(* Logix 5000 project; controller TFF vendor 1 type 14 code 107 rev 33.11; software revision 33.04; part 27 of 38 *)
(* tags used below, declared in another part *)
   Address : DINT;   // Temp Address
   FeedPump_PID_Settings : INT;   // Index
   Index : DINT;   // Index
   TIME : DINT[2];
   AnalogOutput : AnalogOutput[25];   // Analog Output Array
   Concentration : Concentration;
   ControlLoop_FeedPump : ALIAS FOR ControlLoop[1];
   ControlLoop_FeedPumpAlarm : ALIAS FOR AlarmDeviation[1];
   ControlLoop_TIC101 : ALIAS FOR ControlLoop[7];
   DerivedData : DerivedData;   // Derived data (user input and calculated values)
   DF3PHP003 : ALIAS FOR DigitalPoint[27];
   DF48P001 : ALIAS FOR DigitalPoint[23];
   Diafiltration : Diafiltration;
   DigitalOutput : BOOL[256];   // Digital Output Array these bits are sent to output cards.
   DigitalPoint : DigitalPoint[150];   // Digital Point Array
   DP : ALIAS FOR AnalogPoint[40];
   DPAlarm : ALIAS FOR AlarmAnalog[40];
   Drive : Drive[11];   // Drives Array
   FI003 : ALIAS FOR AnalogPoint[42];
   FI101 : ALIAS FOR AnalogPoint[19];
   FI201 : ALIAS FOR AnalogPoint[2];
   FI401 : ALIAS FOR AnalogPoint[20];
   FlowPath : FlowPath[64];   // Flow Path Array
   FQ_Conc : ALIAS FOR Totalizer[0];   // Concentration Totalizer
   FQ_Diaf : ALIAS FOR Totalizer[1];   // DiafiltrationTotalizer
   LI101 : ALIAS FOR AnalogPoint[44];
   Membrane_Data : Membrane_Data;   // Membrane Data
   NWP : ALIAS FOR AnalogPoint[45];
   Options : Options;   // Options List
   PERM : ALIAS FOR AnalogPoint[46];
   Phase0 : ALIAS FOR Phase[0];   // Phase 0
   PI001 : ALIAS FOR AnalogPoint[5];
   PI101 : ALIAS FOR AnalogPoint[6];
   PI201 : ALIAS FOR AnalogPoint[7];
   PipeAnimation : PipeAnimation;   // HMI Pipe Animation Array
   SIC001 : ALIAS FOR Drive[1];
   SIC001DF : ALIAS FOR DigitalPoint[16];
   SIC002 : ALIAS FOR Drive[2];
   SIC003DF : ALIAS FOR DigitalPoint[29];
   SysControl : SysControl;   // General system status and command
   TCU101_AO : ALIAS FOR AnalogOutput[6];
   TI101 : ALIAS FOR AnalogPoint[13];
   TI201 : ALIAS FOR AnalogPoint[22];
   TIC101Control : TCUControl;
   TMP : ALIAS FOR AnalogPoint[41];
   TMPAlarm : ALIAS FOR AlarmAnalog[41];
   XV701 : ALIAS FOR Valve[17];
   XV702 : ALIAS FOR Valve[18];
(* Process, continued *)

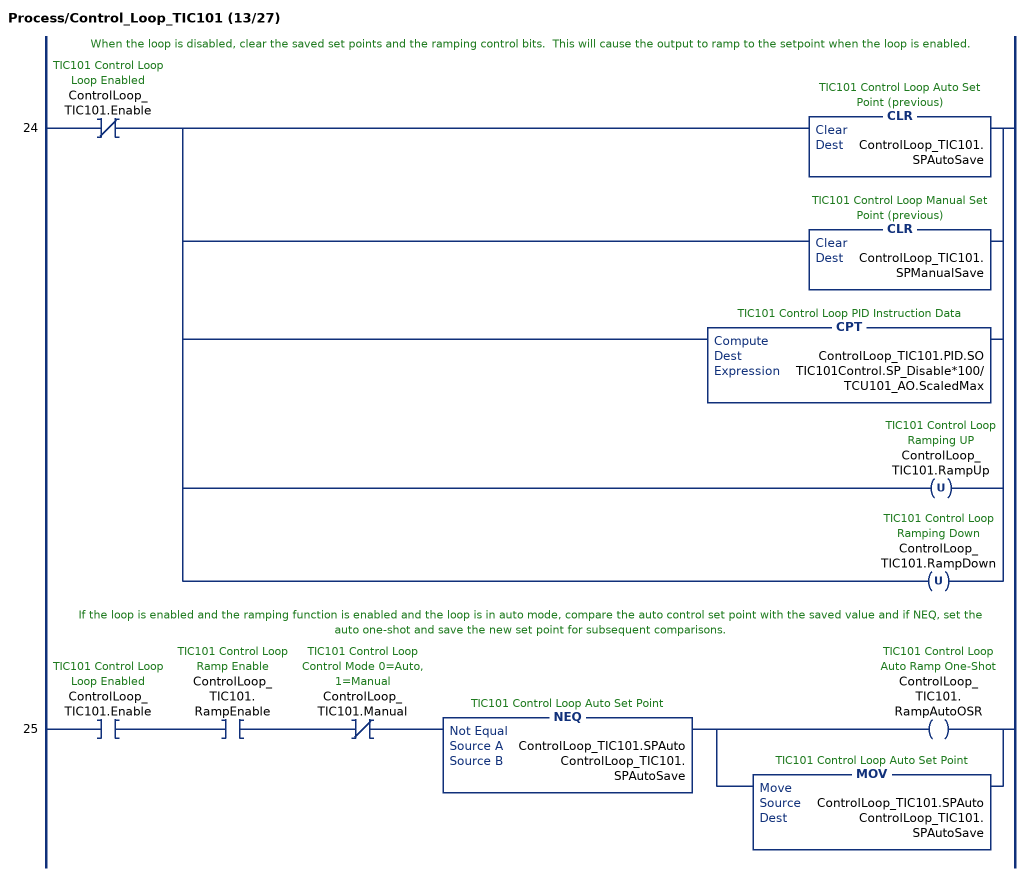
   [picture p263: Process/Control_Loop_TIC101 rungs 24-25]
   // When the loop is disabled, clear the saved set points and the ramping control bits.  This will cause the output to ramp to the setpoint when the loop is enabled.
   24: XIO(ControlLoop_TIC101.Enable)[CLR(ControlLoop_TIC101.SPAutoSave) ,CLR(ControlLoop_TIC101.SPManualSave) ,CPT(ControlLoop_TIC101.PID.SO,TIC101Control.SP_Disable*100/TCU101_AO.ScaledMax) ,OTU(ControlLoop_TIC101.RampUp) ,OTU(ControlLoop_TIC101.RampDown) ];
   // If the loop is enabled and the ramping function is enabled and the loop is in auto mode, compare the auto control set point with the saved value and if NEQ, set the auto one-shot and save the new set point for subsequent comparisons.
   25: XIC(ControlLoop_TIC101.Enable)XIC(ControlLoop_TIC101.RampEnable)XIO(ControlLoop_TIC101.Manual)NEQ(ControlLoop_TIC101.SPAuto,ControlLoop_TIC101.SPAutoSave)[OTE(ControlLoop_TIC101.RampAutoOSR) ,MOV(ControlLoop_TIC101.SPAuto,ControlLoop_TIC101.SPAutoSave) ];
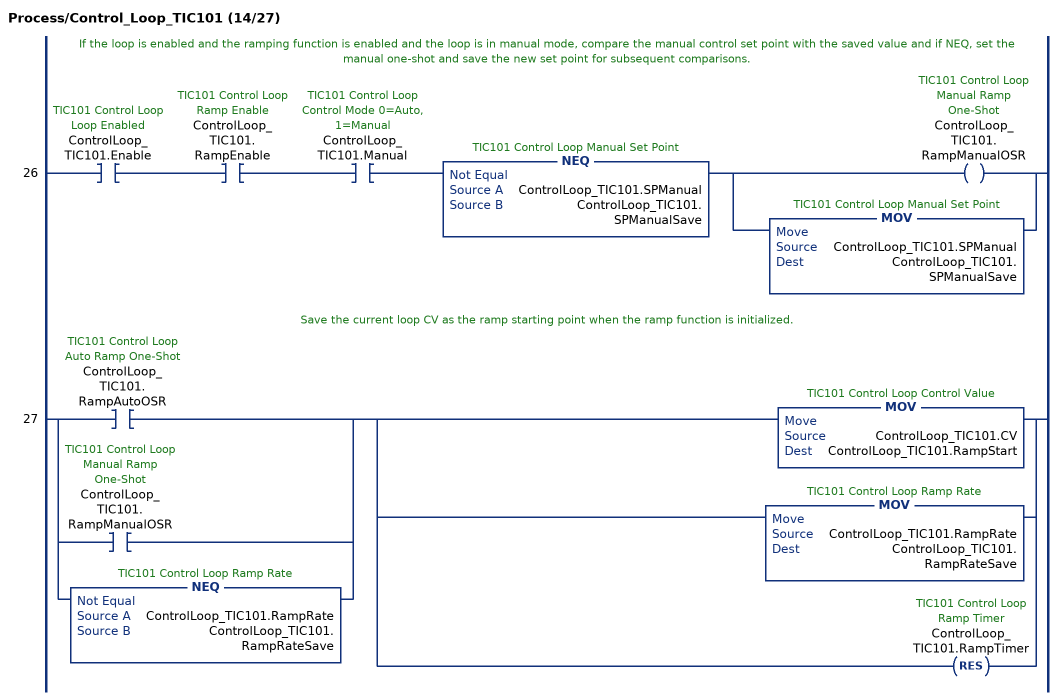
   // If the loop is enabled and the ramping function is enabled and the loop is in manual mode, compare the manual control set point with the saved value and if NEQ, set the manual one-shot and save the new set point for subsequent comparisons.
   26: XIC(ControlLoop_TIC101.Enable)XIC(ControlLoop_TIC101.RampEnable)XIC(ControlLoop_TIC101.Manual)NEQ(ControlLoop_TIC101.SPManual,ControlLoop_TIC101.SPManualSave)[OTE(ControlLoop_TIC101.RampManualOSR) ,MOV(ControlLoop_TIC101.SPManual,ControlLoop_TIC101.SPManualSave) ];
   // Save the current loop CV as the ramp starting point when the ramp function is initialized.
   27: [XIC(ControlLoop_TIC101.RampAutoOSR) ,XIC(ControlLoop_TIC101.RampManualOSR) ,NEQ(ControlLoop_TIC101.RampRate,ControlLoop_TIC101.RampRateSave) ][MOV(ControlLoop_TIC101.CV,ControlLoop_TIC101.RampStart) ,MOV(ControlLoop_TIC101.RampRate,ControlLoop_TIC101.RampRateSave) ,RES(ControlLoop_TIC101.RampTimer) ];
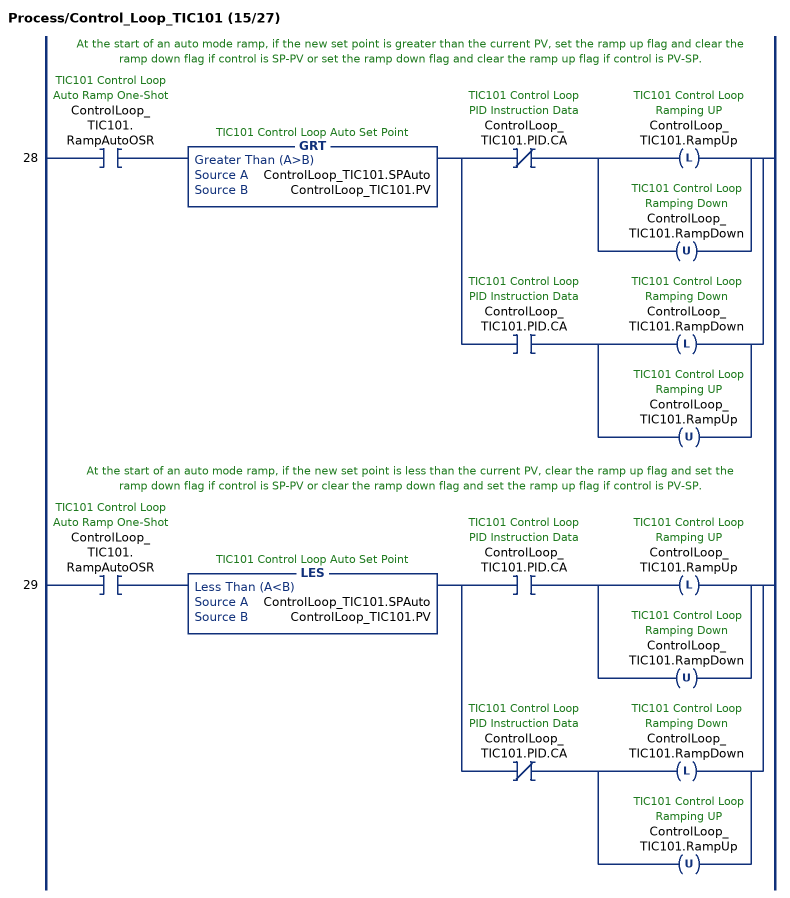
   // At the start of an auto mode ramp, if the new set point is greater than the current PV, set the ramp up flag and clear the ramp down flag if control is SP-PV or set the ramp down flag and clear the ramp up flag if control is PV-SP.
   28: XIC(ControlLoop_TIC101.RampAutoOSR)GRT(ControlLoop_TIC101.SPAuto,ControlLoop_TIC101.PV)[XIO(ControlLoop_TIC101.PID.CA) [OTL(ControlLoop_TIC101.RampUp) ,OTU(ControlLoop_TIC101.RampDown) ] ,XIC(ControlLoop_TIC101.PID.CA) [OTL(ControlLoop_TIC101.RampDown) ,OTU(ControlLoop_TIC101.RampUp) ] ];
   // At the start of an auto mode ramp, if the new set point is less than the current PV, clear the ramp up flag and set the ramp down flag if control is SP-PV or clear the ramp down flag and set the ramp up flag if control is PV-SP.
   29: XIC(ControlLoop_TIC101.RampAutoOSR)LES(ControlLoop_TIC101.SPAuto,ControlLoop_TIC101.PV)[XIC(ControlLoop_TIC101.PID.CA) [OTL(ControlLoop_TIC101.RampUp) ,OTU(ControlLoop_TIC101.RampDown) ] ,XIO(ControlLoop_TIC101.PID.CA) [OTL(ControlLoop_TIC101.RampDown) ,OTU(ControlLoop_TIC101.RampUp) ] ];
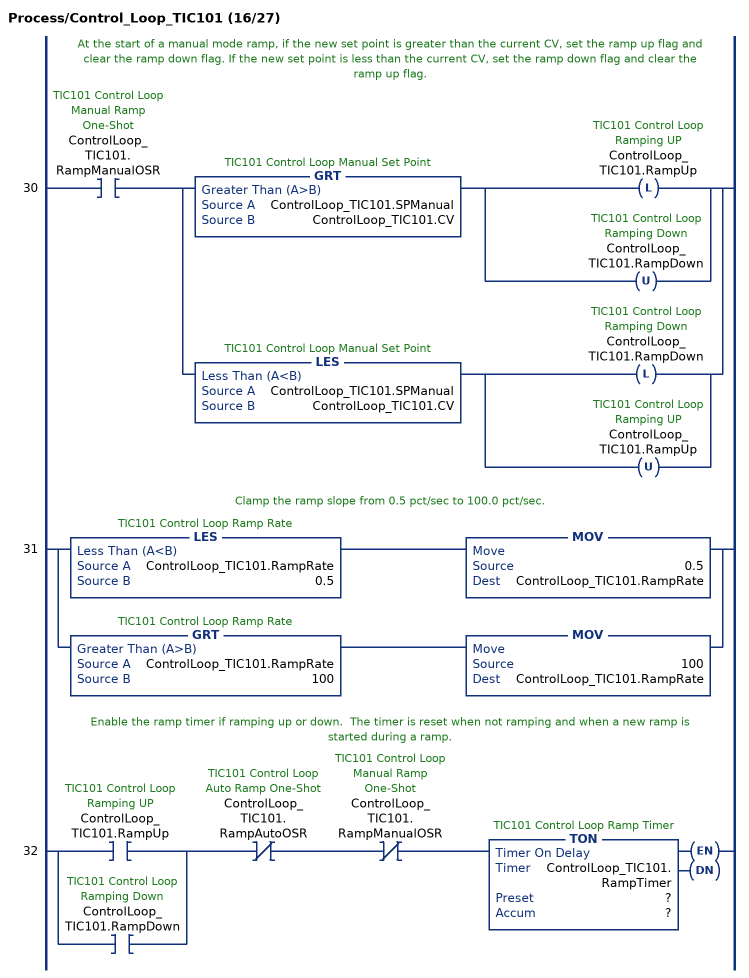
   // At the start of a manual mode ramp, if the new set point is greater than the current CV, set the ramp up flag and clear the ramp down flag. If the new set point is less than the current CV, set the ramp down flag and clear the ramp up flag.
   30: XIC(ControlLoop_TIC101.RampManualOSR)[GRT(ControlLoop_TIC101.SPManual,ControlLoop_TIC101.CV) [OTL(ControlLoop_TIC101.RampUp) ,OTU(ControlLoop_TIC101.RampDown) ] ,LES(ControlLoop_TIC101.SPManual,ControlLoop_TIC101.CV) [OTL(ControlLoop_TIC101.RampDown) ,OTU(ControlLoop_TIC101.RampUp) ] ];
   // Clamp the ramp slope from 0.5 pct/sec to 100.0 pct/sec.
   31: [LES(ControlLoop_TIC101.RampRate,0.5) MOV(0.5,ControlLoop_TIC101.RampRate) ,GRT(ControlLoop_TIC101.RampRate,100) MOV(100,ControlLoop_TIC101.RampRate) ];
   // Enable the ramp timer if ramping up or down.  The timer is reset when not ramping and when a new ramp is started during a ramp.
   32: [XIC(ControlLoop_TIC101.RampUp) ,XIC(ControlLoop_TIC101.RampDown) ]XIO(ControlLoop_TIC101.RampAutoOSR)XIO(ControlLoop_TIC101.RampManualOSR)TON(ControlLoop_TIC101.RampTimer,?,?);
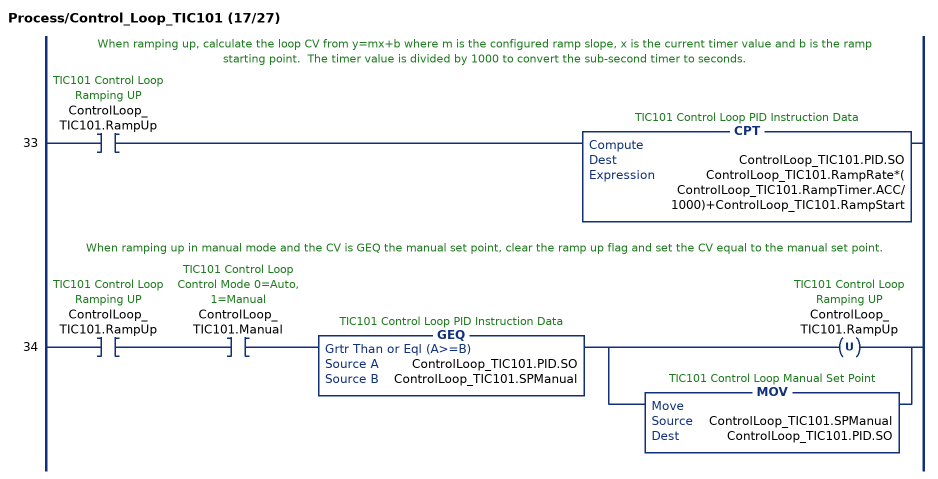
   // When ramping up, calculate the loop CV from y=mx+b where m is the configured ramp slope, x is the current timer value and b is the ramp starting point.  The timer value is divided by 1000 to convert the sub-second timer to seconds.
   33: XIC(ControlLoop_TIC101.RampUp)CPT(ControlLoop_TIC101.PID.SO,ControlLoop_TIC101.RampRate*(ControlLoop_TIC101.RampTimer.ACC/1000)+ControlLoop_TIC101.RampStart);
   // When ramping up in manual mode and the CV is GEQ the manual set point, clear the ramp up flag and set the CV equal to the manual set point.
   34: XIC(ControlLoop_TIC101.RampUp)XIC(ControlLoop_TIC101.Manual)GEQ(ControlLoop_TIC101.PID.SO,ControlLoop_TIC101.SPManual)[OTU(ControlLoop_TIC101.RampUp) ,MOV(ControlLoop_TIC101.SPManual,ControlLoop_TIC101.PID.SO) ];
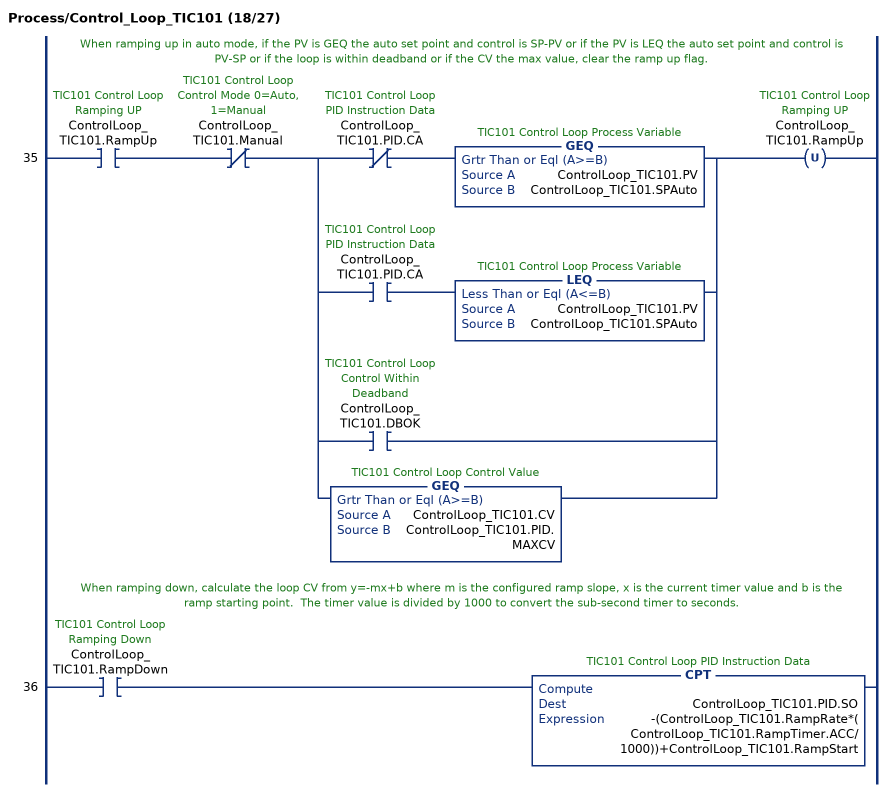
   // When ramping up in auto mode, if the PV is GEQ the auto set point and control is SP-PV or if the PV is LEQ the auto set point and control is PV-SP or if the loop is within deadband or if the CV the max value, clear the ramp up flag.
   35: XIC(ControlLoop_TIC101.RampUp)XIO(ControlLoop_TIC101.Manual)[XIO(ControlLoop_TIC101.PID.CA) GEQ(ControlLoop_TIC101.PV,ControlLoop_TIC101.SPAuto) ,XIC(ControlLoop_TIC101.PID.CA) LEQ(ControlLoop_TIC101.PV,ControlLoop_TIC101.SPAuto) ,XIC(ControlLoop_TIC101.DBOK) ,GEQ(ControlLoop_TIC101.CV,ControlLoop_TIC101.PID.MAXCV) ]OTU(ControlLoop_TIC101.RampUp);
   // When ramping down, calculate the loop CV from y=-mx+b where m is the configured ramp slope, x is the current timer value and b is the ramp starting point.  The timer value is divided by 1000 to convert the sub-second timer to seconds.
   36: XIC(ControlLoop_TIC101.RampDown)CPT(ControlLoop_TIC101.PID.SO,-(ControlLoop_TIC101.RampRate*(ControlLoop_TIC101.RampTimer.ACC/1000))+ControlLoop_TIC101.RampStart);
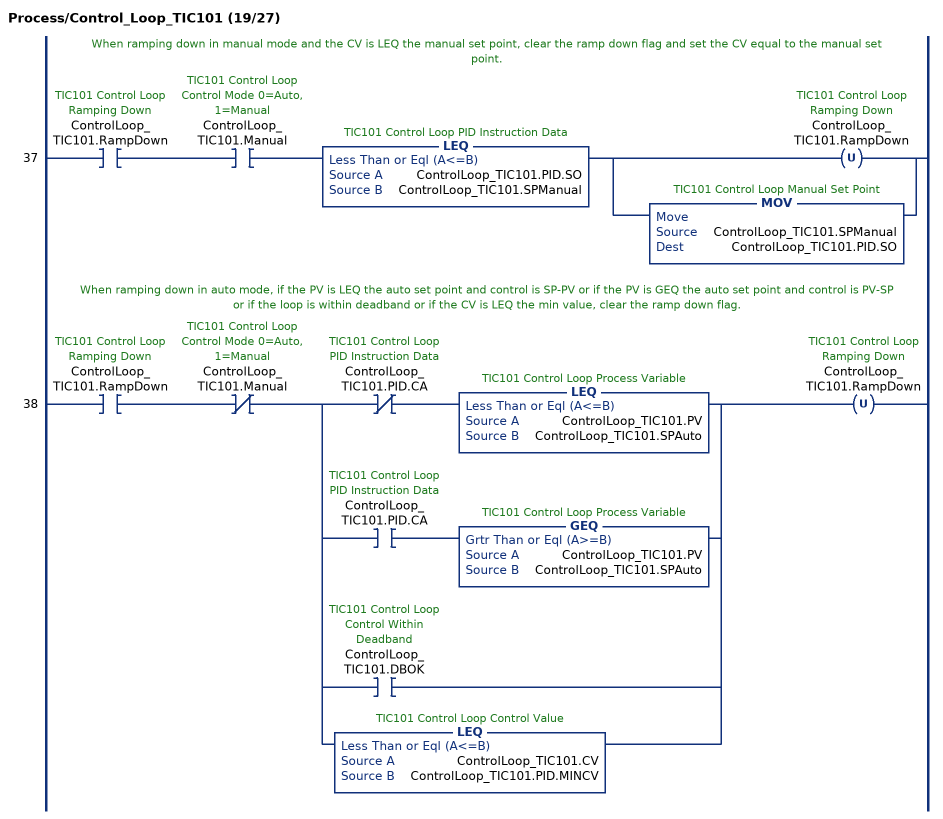
   // When ramping down in manual mode and the CV is LEQ the manual set point, clear the ramp down flag and set the CV equal to the manual set point.
   37: XIC(ControlLoop_TIC101.RampDown)XIC(ControlLoop_TIC101.Manual)LEQ(ControlLoop_TIC101.PID.SO,ControlLoop_TIC101.SPManual)[OTU(ControlLoop_TIC101.RampDown) ,MOV(ControlLoop_TIC101.SPManual,ControlLoop_TIC101.PID.SO) ];
   // When ramping down in auto mode, if the PV is LEQ the auto set point and control is SP-PV or if the PV is GEQ the auto set point and control is PV-SP or if the loop is within deadband or if the CV is LEQ the min value, clear the ramp down flag.
   38: XIC(ControlLoop_TIC101.RampDown)XIO(ControlLoop_TIC101.Manual)[XIO(ControlLoop_TIC101.PID.CA) LEQ(ControlLoop_TIC101.PV,ControlLoop_TIC101.SPAuto) ,XIC(ControlLoop_TIC101.PID.CA) GEQ(ControlLoop_TIC101.PV,ControlLoop_TIC101.SPAuto) ,XIC(ControlLoop_TIC101.DBOK) ,LEQ(ControlLoop_TIC101.CV,ControlLoop_TIC101.PID.MINCV) ]OTU(ControlLoop_TIC101.RampDown);
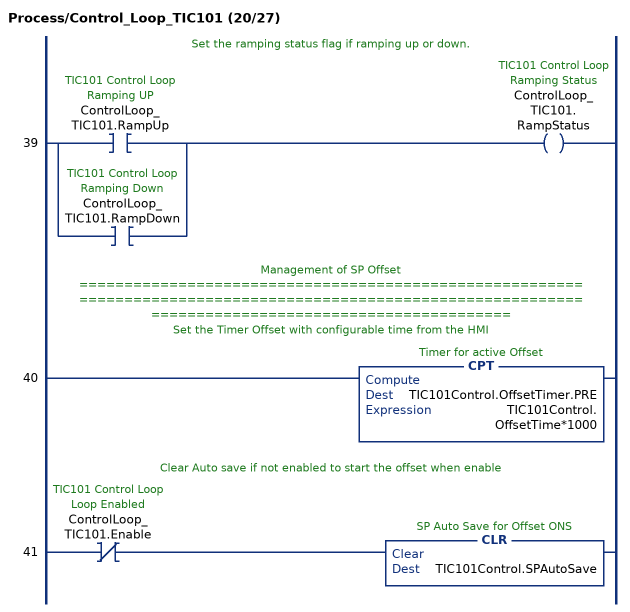
   // Set the ramping status flag if ramping up or down.
   39: [XIC(ControlLoop_TIC101.RampUp) ,XIC(ControlLoop_TIC101.RampDown) ]OTE(ControlLoop_TIC101.RampStatus);
   // Management of SP Offset
   // ========================================================================================================================================================
   // Set the Timer Offset with configurable time from the HMI
   40: CPT(TIC101Control.OffsetTimer.PRE,TIC101Control.OffsetTime*1000);
   // Clear Auto save if not enabled to start the offset when enable
   41: XIO(ControlLoop_TIC101.Enable)CLR(TIC101Control.SPAutoSave);
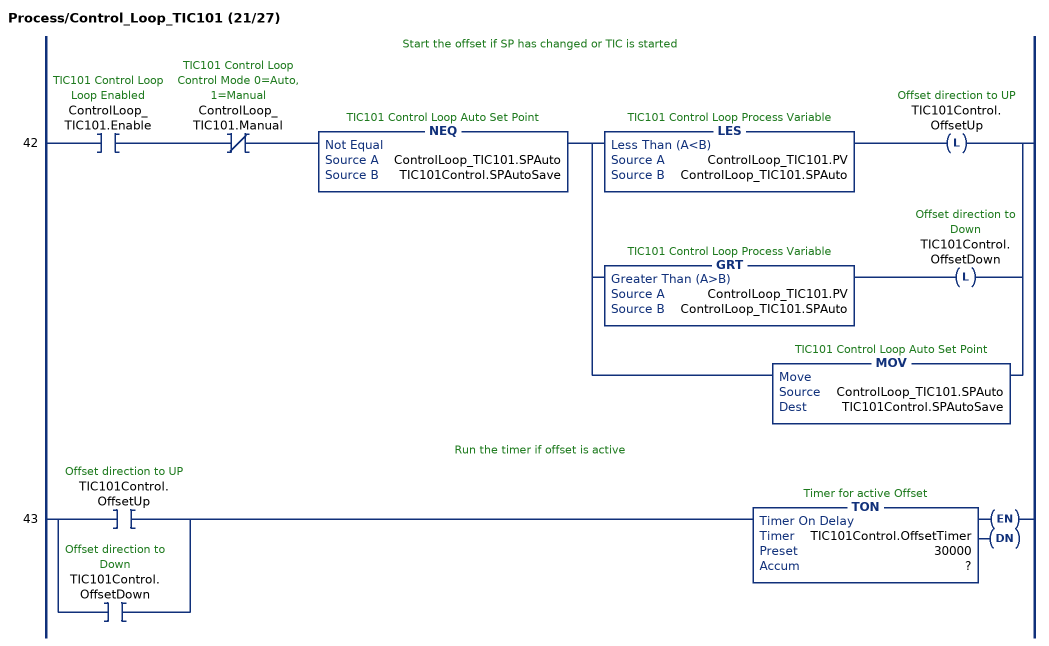
   // Start the offset if SP has changed or TIC is started
   42: XIC(ControlLoop_TIC101.Enable)XIO(ControlLoop_TIC101.Manual)NEQ(ControlLoop_TIC101.SPAuto,TIC101Control.SPAutoSave)[[LES(ControlLoop_TIC101.PV,ControlLoop_TIC101.SPAuto) OTL(TIC101Control.OffsetUp) ,GRT(ControlLoop_TIC101.PV,ControlLoop_TIC101.SPAuto) OTL(TIC101Control.OffsetDown) ] ,MOV(ControlLoop_TIC101.SPAuto,TIC101Control.SPAutoSave) ];
   // Run the timer if offset is active
   43: [XIC(TIC101Control.OffsetUp) ,XIC(TIC101Control.OffsetDown) ]TON(TIC101Control.OffsetTimer,?,?);
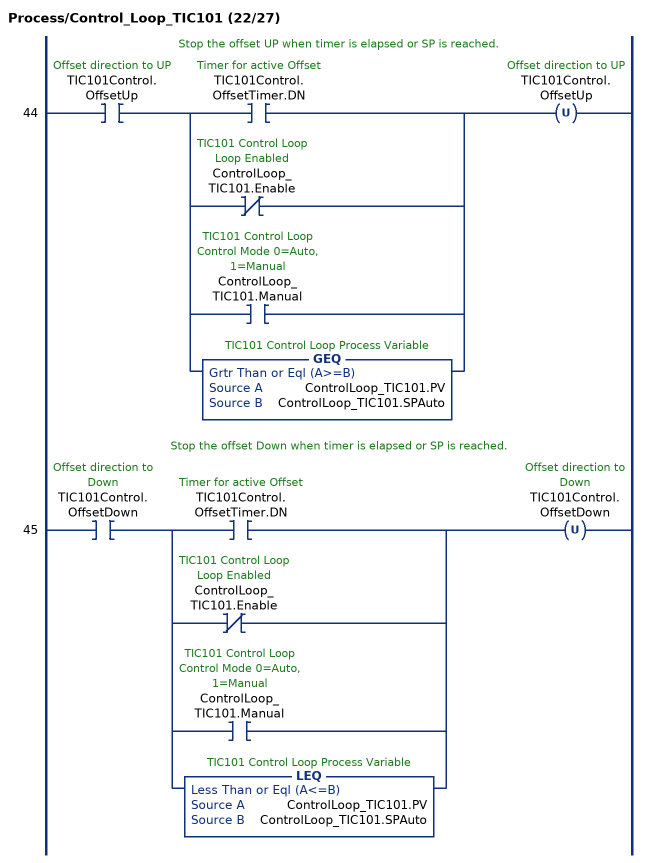
   // Stop the offset UP when timer is elapsed or SP is reached.
   44: XIC(TIC101Control.OffsetUp)[XIC(TIC101Control.OffsetTimer.DN) ,XIO(ControlLoop_TIC101.Enable) ,XIC(ControlLoop_TIC101.Manual) ,GEQ(ControlLoop_TIC101.PV,ControlLoop_TIC101.SPAuto) ]OTU(TIC101Control.OffsetUp);
   // Stop the offset Down when timer is elapsed or SP is reached.
   45: XIC(TIC101Control.OffsetDown)[XIC(TIC101Control.OffsetTimer.DN) ,XIO(ControlLoop_TIC101.Enable) ,XIC(ControlLoop_TIC101.Manual) ,LEQ(ControlLoop_TIC101.PV,ControlLoop_TIC101.SPAuto) ]OTU(TIC101Control.OffsetDown);
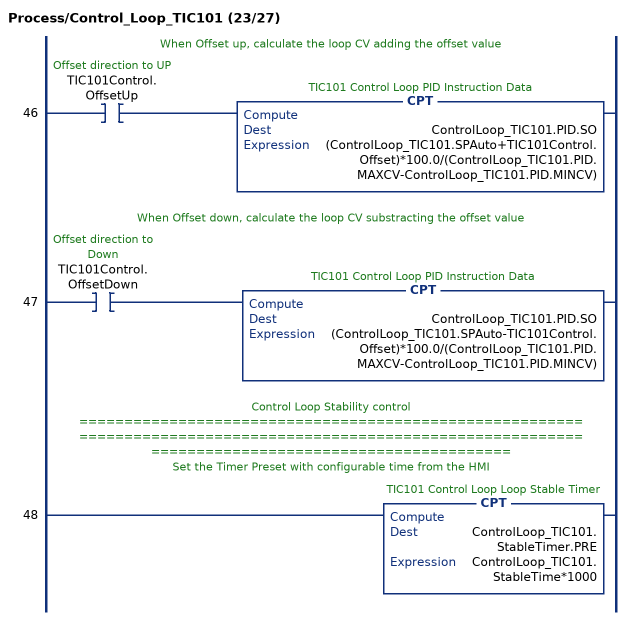
   // When Offset up, calculate the loop CV adding the offset value
   46: XIC(TIC101Control.OffsetUp)CPT(ControlLoop_TIC101.PID.SO,(ControlLoop_TIC101.SPAuto+TIC101Control.Offset)*100.0/(ControlLoop_TIC101.PID.MAXCV-ControlLoop_TIC101.PID.MINCV));
   // When Offset down, calculate the loop CV substracting the offset value
   47: XIC(TIC101Control.OffsetDown)CPT(ControlLoop_TIC101.PID.SO,(ControlLoop_TIC101.SPAuto-TIC101Control.Offset)*100.0/(ControlLoop_TIC101.PID.MAXCV-ControlLoop_TIC101.PID.MINCV));
   // Control Loop Stability control
   // ========================================================================================================================================================
   // Set the Timer Preset with configurable time from the HMI
   48: CPT(ControlLoop_TIC101.StableTimer.PRE,ControlLoop_TIC101.StableTime*1000);
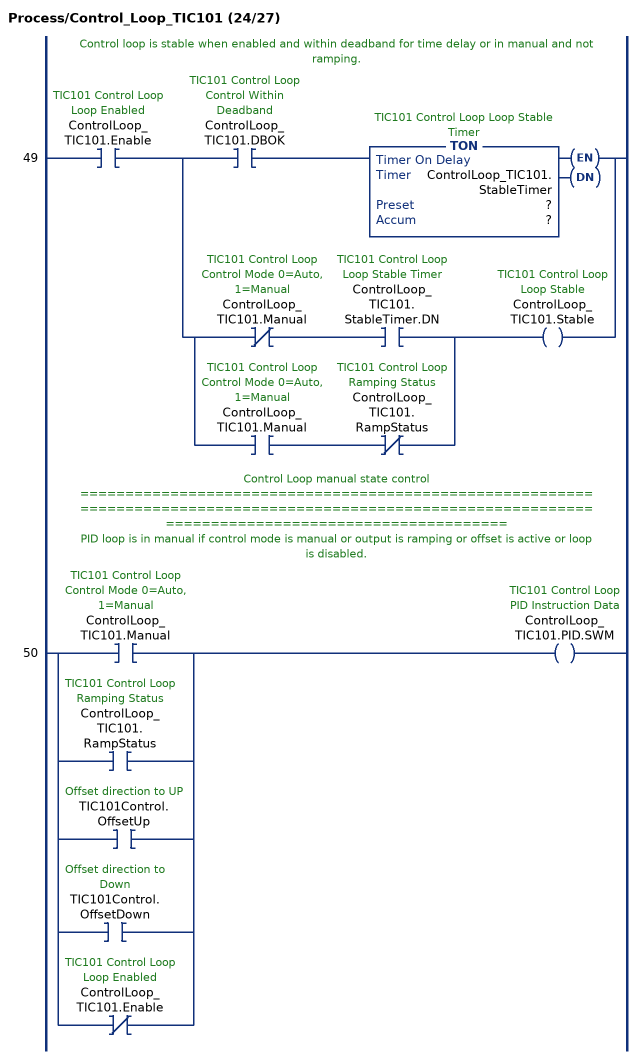
   // Control loop is stable when enabled and within deadband for time delay or in manual and not ramping.
   49: XIC(ControlLoop_TIC101.Enable)[XIC(ControlLoop_TIC101.DBOK) TON(ControlLoop_TIC101.StableTimer,?,?) ,[XIO(ControlLoop_TIC101.Manual) XIC(ControlLoop_TIC101.StableTimer.DN) ,XIC(ControlLoop_TIC101.Manual) XIO(ControlLoop_TIC101.RampStatus) ] OTE(ControlLoop_TIC101.Stable) ];
   // Control Loop manual state control
   // ========================================================================================================================================================
   // PID loop is in manual if control mode is manual or output is ramping or offset is active or loop is disabled.
   50: [XIC(ControlLoop_TIC101.Manual) ,XIC(ControlLoop_TIC101.RampStatus) ,XIC(TIC101Control.OffsetUp) ,XIC(TIC101Control.OffsetDown) ,XIO(ControlLoop_TIC101.Enable) ]OTE(ControlLoop_TIC101.PID.SWM);
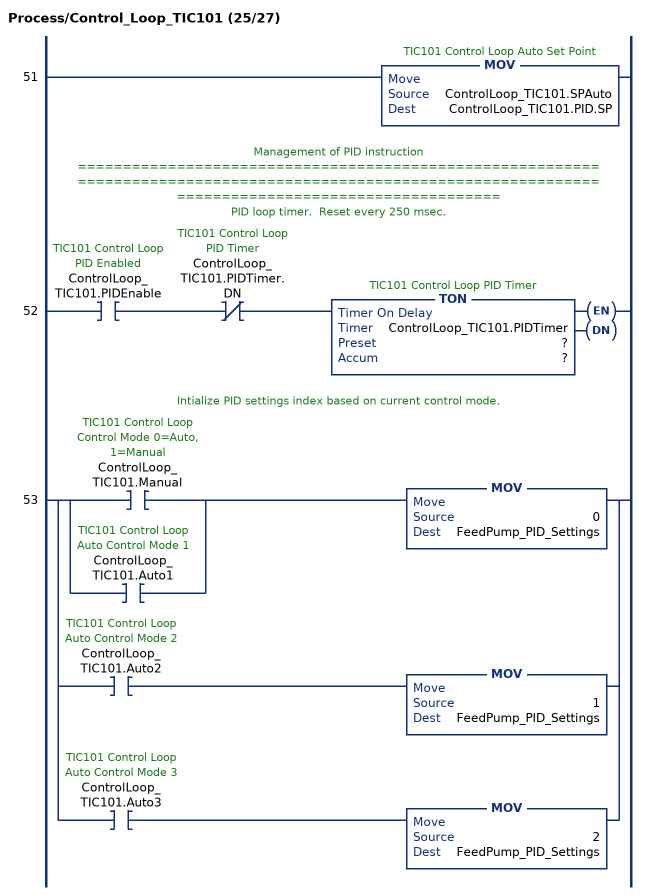
   51: MOV(ControlLoop_TIC101.SPAuto,ControlLoop_TIC101.PID.SP);
   // Management of PID instruction
   // ========================================================================================================================================================
   // PID loop timer.  Reset every 250 msec.
   52: XIC(ControlLoop_TIC101.PIDEnable)XIO(ControlLoop_TIC101.PIDTimer.DN)TON(ControlLoop_TIC101.PIDTimer,?,?);
   // Intialize PID settings index based on current control mode.
   53: [[XIC(ControlLoop_TIC101.Manual) ,XIC(ControlLoop_TIC101.Auto1) ] MOV(0,FeedPump_PID_Settings) ,XIC(ControlLoop_TIC101.Auto2) MOV(1,FeedPump_PID_Settings) ,XIC(ControlLoop_TIC101.Auto3) MOV(2,FeedPump_PID_Settings) ];
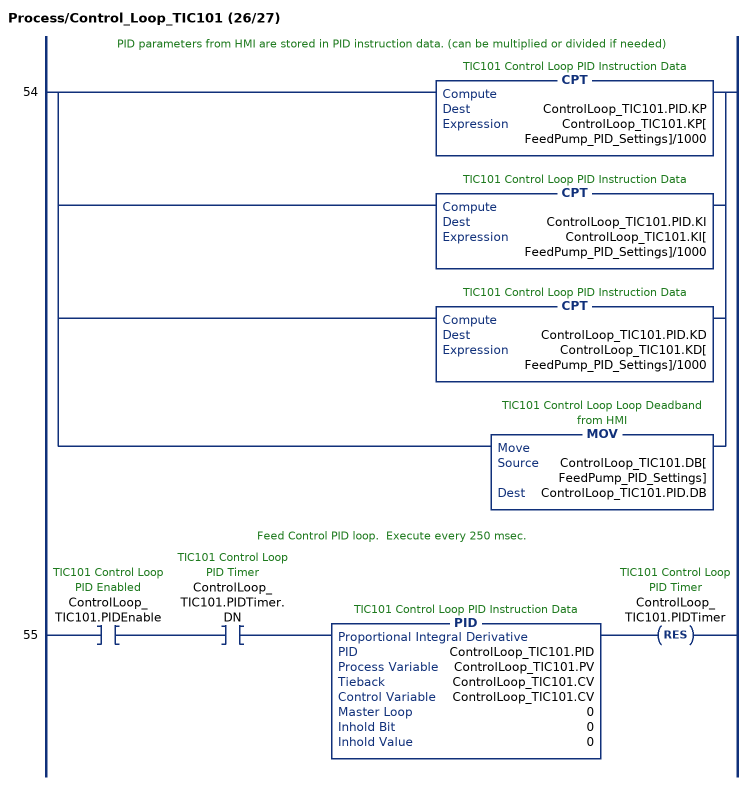
   // PID parameters from HMI are stored in PID instruction data. (can be multiplied or divided if needed)
   54: [CPT(ControlLoop_TIC101.PID.KP,ControlLoop_TIC101.KP[FeedPump_PID_Settings]/1000) ,CPT(ControlLoop_TIC101.PID.KI,ControlLoop_TIC101.KI[FeedPump_PID_Settings]/1000) ,CPT(ControlLoop_TIC101.PID.KD,ControlLoop_TIC101.KD[FeedPump_PID_Settings]/1000) ,MOV(ControlLoop_TIC101.DB[FeedPump_PID_Settings],ControlLoop_TIC101.PID.DB) ];
   // Feed Control PID loop.  Execute every 250 msec.
   55: XIC(ControlLoop_TIC101.PIDEnable)XIC(ControlLoop_TIC101.PIDTimer.DN)PID(ControlLoop_TIC101.PID,ControlLoop_TIC101.PV,ControlLoop_TIC101.CV,ControlLoop_TIC101.CV,0,0,0)RES(ControlLoop_TIC101.PIDTimer);
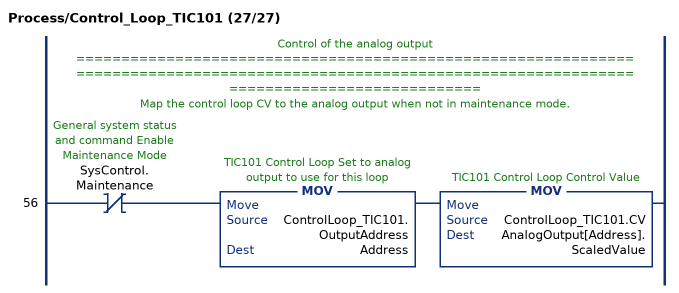
   // Control of the analog output
   // ========================================================================================================================================================
   // Map the control loop CV to the analog output when not in maintenance mode.
   56: XIO(SysControl.Maintenance)MOV(ControlLoop_TIC101.OutputAddress,Address)MOV(ControlLoop_TIC101.CV,AnalogOutput[Address].ScaledValue);
END_ROUTINE

ROUTINE Derived_Data   (* structured text *)
// Derived Data Routine
   (* =======================================================================
   	Derived Data : calculations of derived data
   
   	List of treatments
   		- Derived Data Calculation
   
   -----------------------------------------------------------------------------------------------------------------------------------------------------
   	History
   		2019-DEC-24 - Merck - Q. Spindler - Initial version for Candidate Release 1.00.00.00.a
   		2021-APR-20 - Merck - Q. Spindler - Modifications for Candidate Release 1.00.00.00.e
   					- Add FiltrateUltrasonicFlow option for FI201 Qmax and K factor calculation
   		2022-SEP-23 - Actemium - J. Jaekel - Modifications for Candidate Release 1.01.00.01.a
   					- Use TI201 for NWP when FiltrateCondPH or FiltrateCondPHUV option is enable
   =============================================================================================================================*)
   
   
   (* Derived Data Calculation
   =============================================================================================================================*)
   
   (*Flow Calculation : Use Qmax and K factor to calculate Flow current value*)
   IF NOT(SysControl.Simulate) THEN
   	FI101.CurrentValue := ((FI101.FilteredRaw - FI101.RawMin) / (FI101.RawMax - FI101.RawMin)) * DerivedData.FI101Q * DerivedData.FI101K;
   	IF NOT(Options.FiltrateUltrasonicFlow) THEN
   		FI201.CurrentValue := ((FI201.FilteredRaw - FI201.RawMin) / (FI201.RawMax - FI201.RawMin)) * DerivedData.FI201Q * DerivedData.FI201K;
   	END_IF;
   	FI401.CurrentValue := ((FI401.FilteredRaw - FI401.RawMin) / (FI401.RawMax - FI401.RawMin)) * DerivedData.FI401Q * DerivedData.FI401K;
   END_IF;
   
   (*If pumps are off or flow is negative set flow to zero *)
   IF NOT SysControl.Simulate THEN
   	IF NOT(SIC001.RunCommand) OR FI101.CurrentValue < 0 THEN FI101.CurrentValue := 0; END_IF;
   	IF NOT(SIC001.RunCommand) OR FI201.CurrentValue < 0 THEN FI201.CurrentValue := 0; END_IF;
   	IF NOT(SIC002.RunCommand) OR FI401.CurrentValue < 0 THEN FI401.CurrentValue := 0; END_IF;
   END_IF;
   
   (* Feed Flow Calculation*)
   FI003.CurrentValue := (FI101.CurrentValue + FI201.CurrentValue);
   
   
   (*Differential Pressure*)
   DP.CurrentValue := PI001.CurrentValue - PI101.CurrentValue;
   DPAlarm.PV := DP.CurrentValue;
   
   
   (*Trans-Membrane Pressure*)
   TMP.CurrentValue := ((PI001.CurrentValue + PI101.CurrentValue) / 2) - PI201.CurrentValue;
   TMPAlarm.PV := TMP.CurrentValue;
   
   
   (*Flux : Membrane Flux*)
   Membrane_Data.Flux := FI201.CurrentValue / Membrane_Data.Area * 60;
   
   (*Diafiltration Volumes*)
   Diafiltration.Diaf_Volume := FQ_Diaf.Total / (Diafiltration.Diaf_Init + DerivedData.HOLDUP);
   
   (*VCF : Volume Concentration Factor*)
   Concentration.VCF := (LI101.CurrentValue + FQ_Conc.Total) / (LI101.CurrentValue + DerivedData.HOLDUP);
   
   (*Clamp VCF Value if less than 1*)
   IF Concentration.VCF < 1 THEN Concentration.VCF := 1; END_IF;
   
   (*CB : Protein Concentration*)
   Concentration.CB := Concentration.Conc_Init * Concentration.VCF;
   
   
   (*NWP TCF*)
   
   (*Fill Lookup Table for TCF 25 DegC*)
   Membrane_Data.NWP_TCF_Lookup_25[0] := 2.011;
   Membrane_Data.NWP_TCF_Lookup_25[1] := 1.943;
   Membrane_Data.NWP_TCF_Lookup_25[2] := 1.879;
   Membrane_Data.NWP_TCF_Lookup_25[3] := 1.818;
   Membrane_Data.NWP_TCF_Lookup_25[4] := 1.761;
   Membrane_Data.NWP_TCF_Lookup_25[5] := 1.706;
   Membrane_Data.NWP_TCF_Lookup_25[6] := 1.653;
   Membrane_Data.NWP_TCF_Lookup_25[7] := 1.604;
   Membrane_Data.NWP_TCF_Lookup_25[8] := 1.556;
   Membrane_Data.NWP_TCF_Lookup_25[9] := 1.511;
   Membrane_Data.NWP_TCF_Lookup_25[10] := 1.468;
   Membrane_Data.NWP_TCF_Lookup_25[11] := 1.426;
   Membrane_Data.NWP_TCF_Lookup_25[12] := 1.387;
   Membrane_Data.NWP_TCF_Lookup_25[13] := 1.349;
   Membrane_Data.NWP_TCF_Lookup_25[14] := 1.313;
   Membrane_Data.NWP_TCF_Lookup_25[15] := 1.278;
   Membrane_Data.NWP_TCF_Lookup_25[16] := 1.245;
   Membrane_Data.NWP_TCF_Lookup_25[17] := 1.213;
   Membrane_Data.NWP_TCF_Lookup_25[18] := 1.183;
   Membrane_Data.NWP_TCF_Lookup_25[19] := 1.154;
   Membrane_Data.NWP_TCF_Lookup_25[20] := 1.126;
   Membrane_Data.NWP_TCF_Lookup_25[21] := 1.099;
   Membrane_Data.NWP_TCF_Lookup_25[22] := 1.072;
   Membrane_Data.NWP_TCF_Lookup_25[23] := 1.047;
   Membrane_Data.NWP_TCF_Lookup_25[24] := 1.022;
   Membrane_Data.NWP_TCF_Lookup_25[25] := 1.0;
   Membrane_Data.NWP_TCF_Lookup_25[26] := 0.978;
   Membrane_Data.NWP_TCF_Lookup_25[27] := 0.956;
   Membrane_Data.NWP_TCF_Lookup_25[28] := 0.935;
   Membrane_Data.NWP_TCF_Lookup_25[29] := 0.915;
   Membrane_Data.NWP_TCF_Lookup_25[30] := 0.896;
   Membrane_Data.NWP_TCF_Lookup_25[31] := 0.877;
   Membrane_Data.NWP_TCF_Lookup_25[32] := 0.859;
   Membrane_Data.NWP_TCF_Lookup_25[33] := 0.841;
   Membrane_Data.NWP_TCF_Lookup_25[34] := 0.824;
   Membrane_Data.NWP_TCF_Lookup_25[35] := 0.808;
   Membrane_Data.NWP_TCF_Lookup_25[36] := 0.791;
   Membrane_Data.NWP_TCF_Lookup_25[37] := 0.777;
   Membrane_Data.NWP_TCF_Lookup_25[38] := 0.761;
   Membrane_Data.NWP_TCF_Lookup_25[39] := 0.747;
   Membrane_Data.NWP_TCF_Lookup_25[40] := 0.733;
   Membrane_Data.NWP_TCF_Lookup_25[41] := 0.719;
   Membrane_Data.NWP_TCF_Lookup_25[42] := 0.706;
   Membrane_Data.NWP_TCF_Lookup_25[43] := 0.694;
   Membrane_Data.NWP_TCF_Lookup_25[44] := 0.681;
   Membrane_Data.NWP_TCF_Lookup_25[45] := 0.669;
   Membrane_Data.NWP_TCF_Lookup_25[46] := 0.658;
   Membrane_Data.NWP_TCF_Lookup_25[47] := 0.646;
   Membrane_Data.NWP_TCF_Lookup_25[48] := 0.635;
   Membrane_Data.NWP_TCF_Lookup_25[49] := 0.624;
   Membrane_Data.NWP_TCF_Lookup_25[50] := 0.614;
   Membrane_Data.NWP_TCF_Lookup_25[51] := 0.604;
   Membrane_Data.NWP_TCF_Lookup_25[52] := 0.594;
   
   
   if Options.FiltrateCondPH OR Options.FiltrateCondPHUV then
   
   	(*Compute NWP_TCF based on Lookup Table for TCF 25 DegC*)
   	IF TI201.CurrentValue < 0 THEN;
   		(*Temperature below lookup table values*)
   		Membrane_Data.NWP_TCF:= Membrane_Data.NWP_TCF_Lookup_25[0];
   	ELSIF TI201.CurrentValue> 51 THEN;
   		(*Temperature above lookup table values*)
   		Membrane_Data.NWP_TCF:= Membrane_Data.NWP_TCF_Lookup_25[52];
   	ELSE
   		(*Temperature within lookup table values*)
   		Membrane_Data.NWP_TCF_Temp:= TRUNC(TI201.CurrentValue);
   		Membrane_Data.NWP_TCF:= (TI201.CurrentValue-Membrane_Data.NWP_TCF_Temp) * ( Membrane_Data.NWP_TCF_Lookup_25[Membrane_Data.NWP_TCF_Temp+1] - Membrane_Data.NWP_TCF_Lookup_25[Membrane_Data.NWP_TCF_Temp] ) + Membrane_Data.NWP_TCF_Lookup_25[Membrane_Data.NWP_TCF_Temp];
   	END_IF;
   
   else
   
   	(*Compute NWP_TCF based on Lookup Table for TCF 25 DegC*)
   	IF TI101.CurrentValue < 0 THEN;
   		(*Temperature below lookup table values*)
   		Membrane_Data.NWP_TCF:= Membrane_Data.NWP_TCF_Lookup_25[0];
   	ELSIF TI101.CurrentValue> 51 THEN;
   		(*Temperature above lookup table values*)
   		Membrane_Data.NWP_TCF:= Membrane_Data.NWP_TCF_Lookup_25[52];
   	ELSE
   		(*Temperature within lookup table values*)
   		Membrane_Data.NWP_TCF_Temp:= TRUNC(TI101.CurrentValue);
   		Membrane_Data.NWP_TCF:= (TI101.CurrentValue-Membrane_Data.NWP_TCF_Temp) * ( Membrane_Data.NWP_TCF_Lookup_25[Membrane_Data.NWP_TCF_Temp+1] - Membrane_Data.NWP_TCF_Lookup_25[Membrane_Data.NWP_TCF_Temp] ) + Membrane_Data.NWP_TCF_Lookup_25[Membrane_Data.NWP_TCF_Temp];
   	END_IF;
   
   END_IF;
   
   
   (*NWP : Normalized Water Permeability*)
   IF TMP.CurrentValue <> 0 THEN NWP.CurrentValue := Membrane_Data.Flux * Membrane_Data.NWP_TCF / TMP.CurrentValue; ELSE NWP.CurrentValue := 0; END_IF;
   
   (*PERM : Membrane Permeability*)
   IF TMP.CurrentValue <> 0 THEN PERM.CurrentValue := Membrane_Data.Flux / TMP.CurrentValue; ELSE PERM.CurrentValue := 0; END_IF;
   
END_ROUTINE

ROUTINE Drive_SIC001_Feed   (* ladder *)
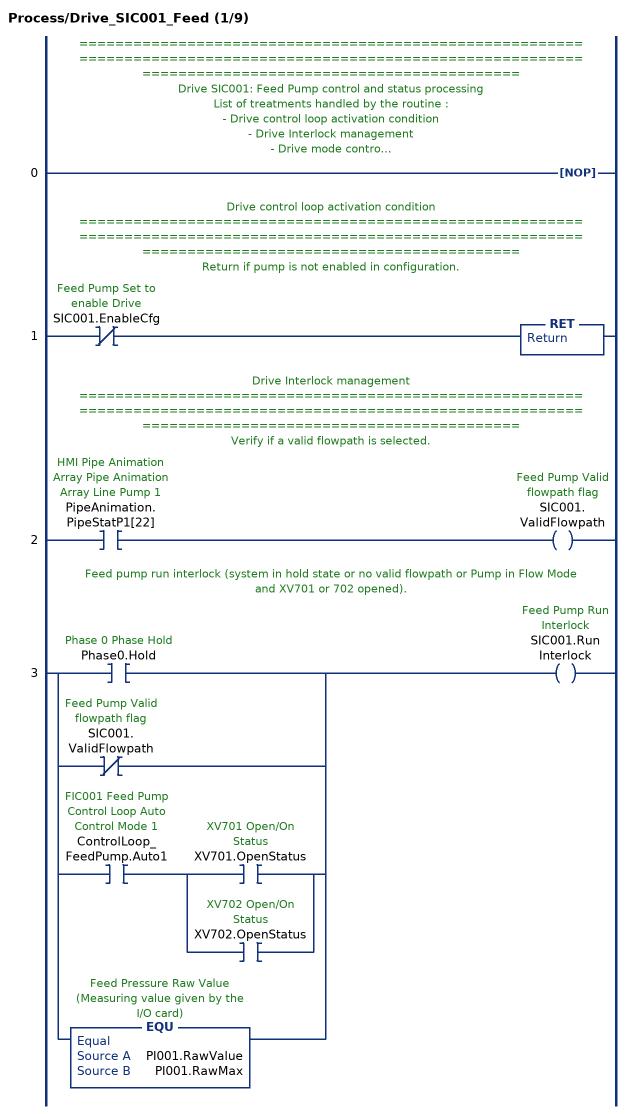
   // ==========================================================================================================================================================
   //                                                    Drive SIC001: Feed Pump control and status processing
   //                                                     List of treatments handled by the routine :
   //                                                          - Drive control loop activation condition
   //                                                          - Drive Interlock management
   //                                                          - Drive mode control
   //                                                          - Drive run command control
   //                                                          - Drive status management
   //                                                          - Drive status for HMI
   //                                                          - Drive DigitalOutput control
   //                                                     -----------------------------------------------------------------------------------------------------------------------------------------------------
   //                                                     History
   // 		2019-DEC-24 - Merck - Q. Spindler - Initial version for Candidate Release 1.00.00.00.a
   // 		2020-APR-06 - Merck - Q. Spindler - Modifications for Candidate Release 1.00.00.00.b
   //                                                                  - Add interlock when XV701 or XV702 is opened and the pump is in flow mode
   //                                                                     - Add interlock when PI001 raw value is equal to RawMax (Sensor disconected)
   // ==========================================================================================================================================================
   0: NOP();
   // Drive control loop activation condition
   // ==========================================================================================================================================================
   // Return if pump is not enabled in configuration.
   1: XIO(SIC001.EnableCfg)RET();
   // Drive Interlock management
   // ==========================================================================================================================================================
   // Verify if a valid flowpath is selected.
   2: XIC(PipeAnimation.PipeStatP1[22])OTE(SIC001.ValidFlowpath);
   // Feed pump run interlock (system in hold state or no valid flowpath or Pump in Flow Mode and XV701 or 702 opened).
   3: [XIC(Phase0.Hold) ,XIO(SIC001.ValidFlowpath) ,XIC(ControlLoop_FeedPump.Auto1) [XIC(XV701.OpenStatus) ,XIC(XV702.OpenStatus) ] ,EQU(PI001.RawValue,PI001.RawMax) ]OTE(SIC001.RunInterlock);
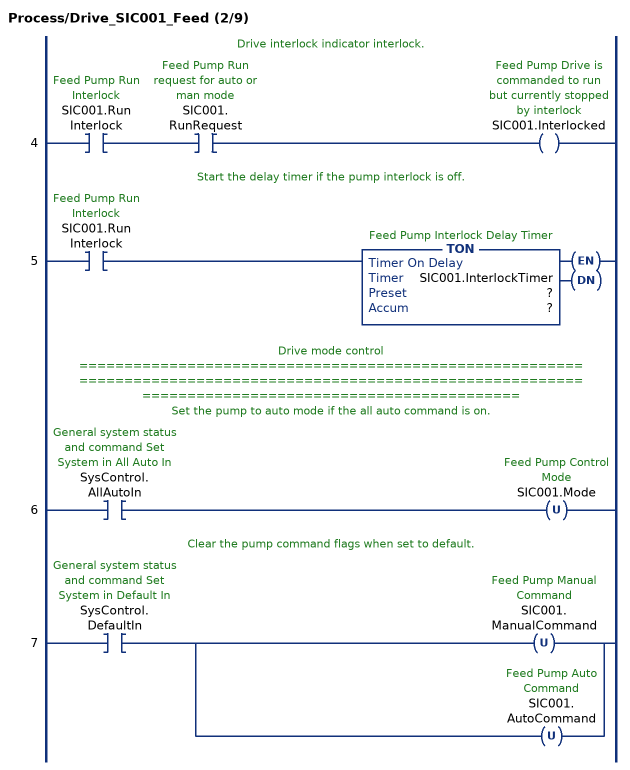
   // Drive interlock indicator interlock.
   4: XIC(SIC001.RunInterlock)XIC(SIC001.RunRequest)OTE(SIC001.Interlocked);
   // Start the delay timer if the pump interlock is off.
   5: XIC(SIC001.RunInterlock)TON(SIC001.InterlockTimer,?,?);
   // Drive mode control
   // ==========================================================================================================================================================
   // Set the pump to auto mode if the all auto command is on.
   6: XIC(SysControl.AllAutoIn)OTU(SIC001.Mode);
   // Clear the pump command flags when set to default.
   7: XIC(SysControl.DefaultIn)[OTU(SIC001.ManualCommand) ,OTU(SIC001.AutoCommand) ];
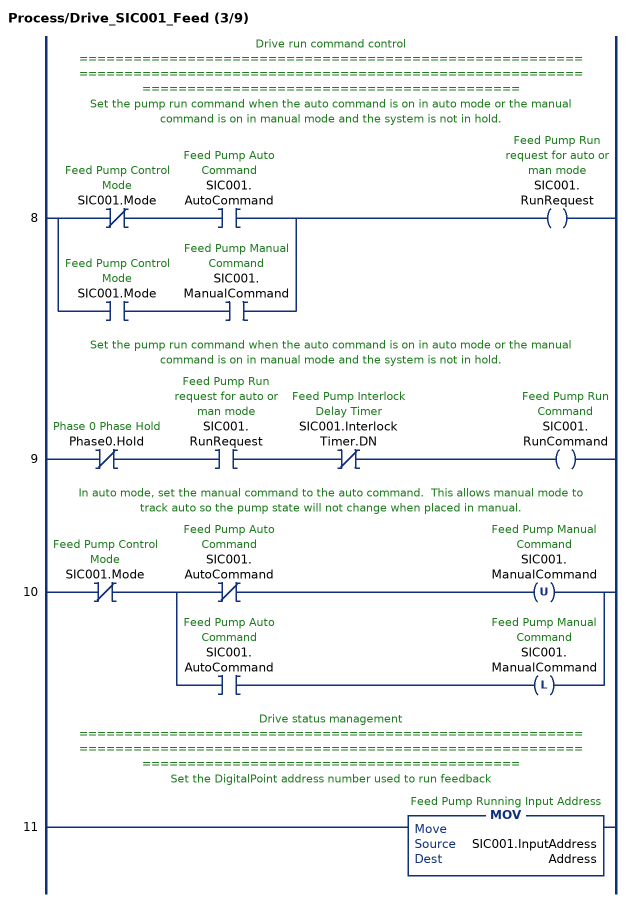
   // Drive run command control
   // ==========================================================================================================================================================
   // Set the pump run command when the auto command is on in auto mode or the manual command is on in manual mode and the system is not in hold.
   8: [XIO(SIC001.Mode) XIC(SIC001.AutoCommand) ,XIC(SIC001.Mode) XIC(SIC001.ManualCommand) ]OTE(SIC001.RunRequest);
   // Set the pump run command when the auto command is on in auto mode or the manual command is on in manual mode and the system is not in hold.
   9: XIO(Phase0.Hold)XIC(SIC001.RunRequest)XIO(SIC001.InterlockTimer.DN)OTE(SIC001.RunCommand);
   // In auto mode, set the manual command to the auto command.  This allows manual mode to track auto so the pump state will not change when placed in manual.
   10: XIO(SIC001.Mode)[XIO(SIC001.AutoCommand) OTU(SIC001.ManualCommand) ,XIC(SIC001.AutoCommand) OTL(SIC001.ManualCommand) ];
   // Drive status management
   // ==========================================================================================================================================================
   // Set the DigitalPoint address number used to run feedback
   11: MOV(SIC001.InputAddress,Address);
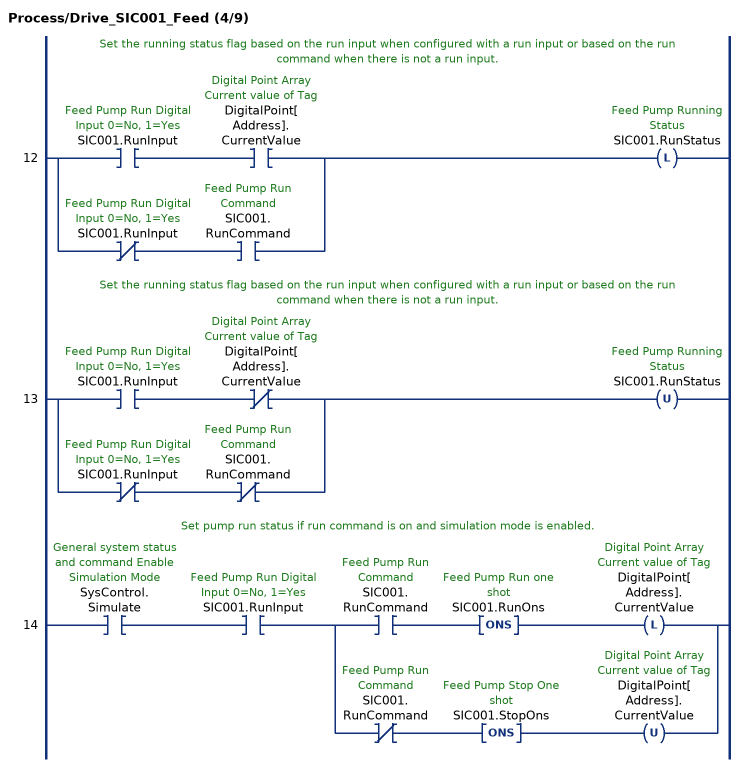
   // Set the running status flag based on the run input when configured with a run input or based on the run command when there is not a run input.
   12: [XIC(SIC001.RunInput) XIC(DigitalPoint[Address].CurrentValue) ,XIO(SIC001.RunInput) XIC(SIC001.RunCommand) ]OTL(SIC001.RunStatus);
   // Set the running status flag based on the run input when configured with a run input or based on the run command when there is not a run input.
   13: [XIC(SIC001.RunInput) XIO(DigitalPoint[Address].CurrentValue) ,XIO(SIC001.RunInput) XIO(SIC001.RunCommand) ]OTU(SIC001.RunStatus);
   // Set pump run status if run command is on and simulation mode is enabled.
   14: XIC(SysControl.Simulate)XIC(SIC001.RunInput)[XIC(SIC001.RunCommand) ONS(SIC001.RunOns) OTL(DigitalPoint[Address].CurrentValue) ,XIO(SIC001.RunCommand) ONS(SIC001.StopOns) OTU(DigitalPoint[Address].CurrentValue) ];
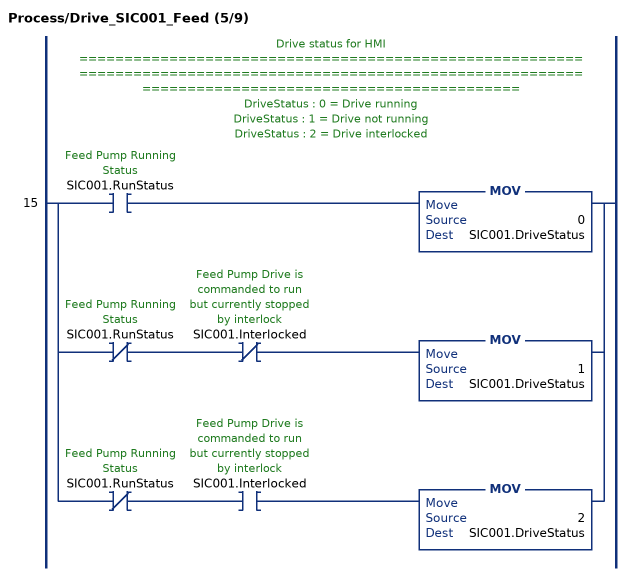
   // Drive status for HMI
   // ==========================================================================================================================================================
   //  DriveStatus : 0 = Drive running
   //  DriveStatus : 1 = Drive not running
   //  DriveStatus : 2 = Drive interlocked
   15: [XIC(SIC001.RunStatus) MOV(0,SIC001.DriveStatus) ,XIO(SIC001.RunStatus) XIO(SIC001.Interlocked) MOV(1,SIC001.DriveStatus) ,XIO(SIC001.RunStatus) XIC(SIC001.Interlocked) MOV(2,SIC001.DriveStatus) ];
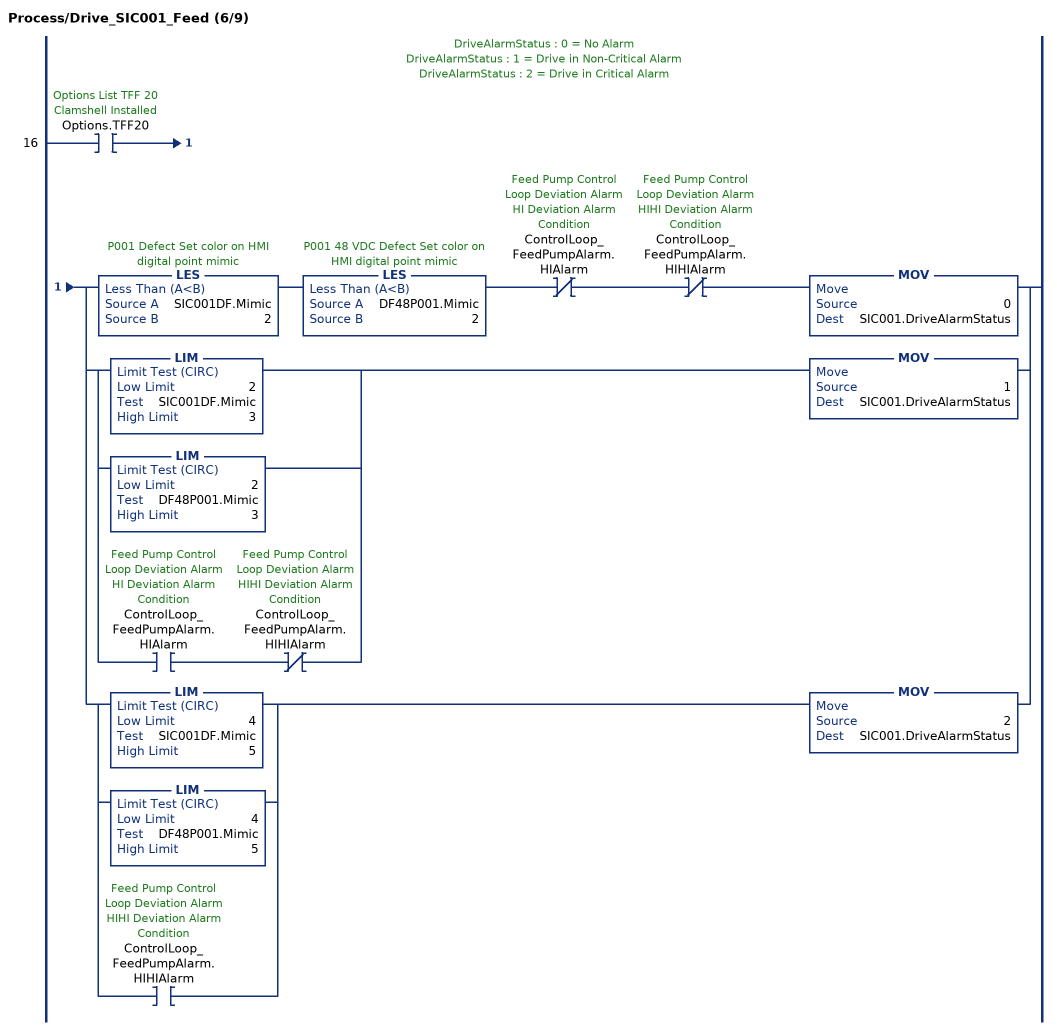
   // DriveAlarmStatus : 0 = No Alarm
   //  DriveAlarmStatus : 1 = Drive in Non-Critical Alarm
   //  DriveAlarmStatus : 2 = Drive in Critical Alarm
   16: XIC(Options.TFF20)[LES(SIC001DF.Mimic,2) LES(DF48P001.Mimic,2) XIO(ControlLoop_FeedPumpAlarm.HIAlarm) XIO(ControlLoop_FeedPumpAlarm.HIHIAlarm) MOV(0,SIC001.DriveAlarmStatus) ,[LIM(2,SIC001DF.Mimic,3) ,LIM(2,DF48P001.Mimic,3) ,XIC(ControlLoop_FeedPumpAlarm.HIAlarm) XIO(ControlLoop_FeedPumpAlarm.HIHIAlarm) ] MOV(1,SIC001.DriveAlarmStatus) ,[LIM(4,SIC001DF.Mimic,5) ,LIM(4,DF48P001.Mimic,5) ,XIC(ControlLoop_FeedPumpAlarm.HIHIAlarm) ] MOV(2,SIC001.DriveAlarmStatus) ];
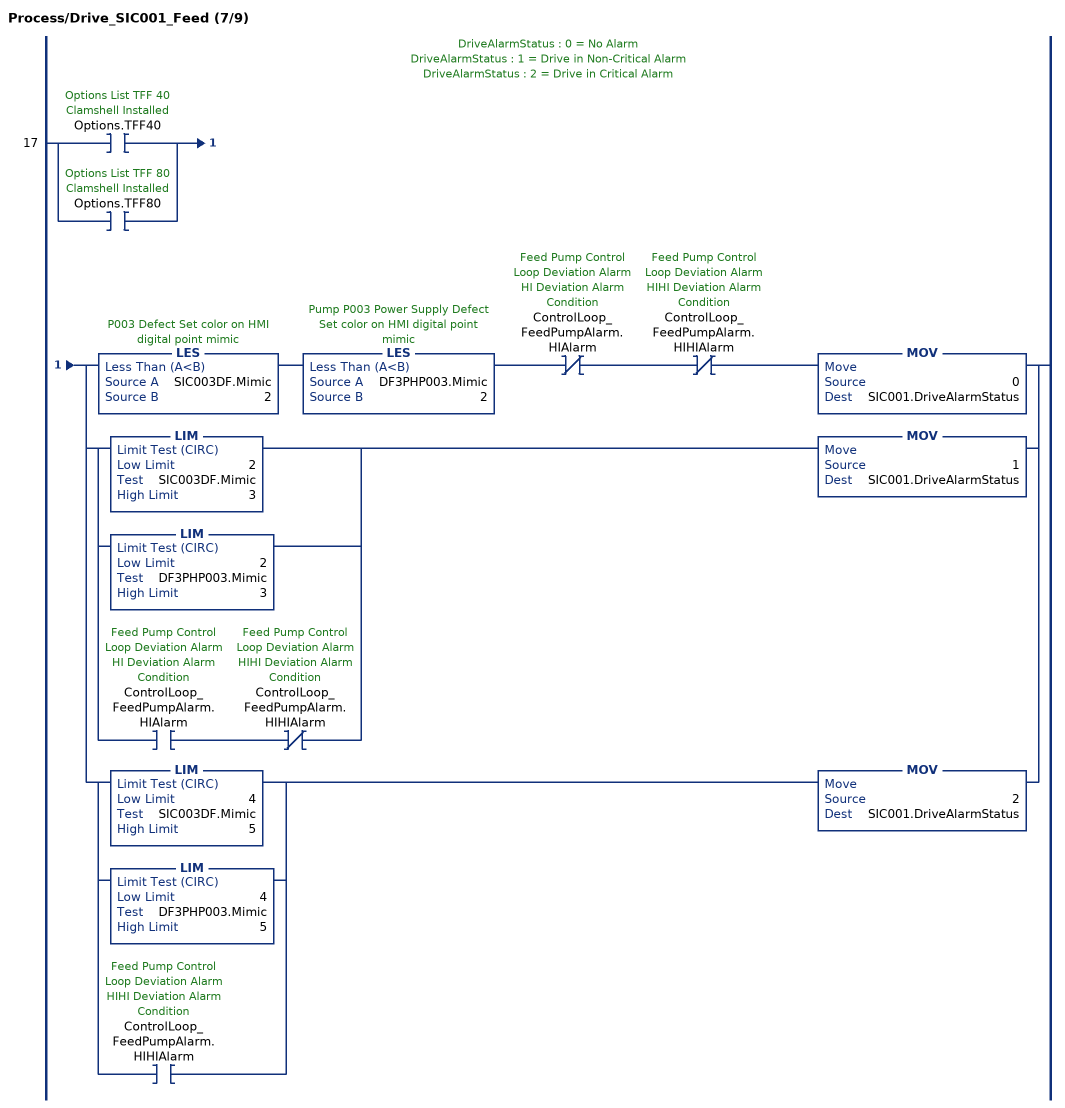
   // DriveAlarmStatus : 0 = No Alarm
   //  DriveAlarmStatus : 1 = Drive in Non-Critical Alarm
   //  DriveAlarmStatus : 2 = Drive in Critical Alarm
   17: [XIC(Options.TFF40) ,XIC(Options.TFF80) ][LES(SIC003DF.Mimic,2) LES(DF3PHP003.Mimic,2) XIO(ControlLoop_FeedPumpAlarm.HIAlarm) XIO(ControlLoop_FeedPumpAlarm.HIHIAlarm) MOV(0,SIC001.DriveAlarmStatus) ,[LIM(2,SIC003DF.Mimic,3) ,LIM(2,DF3PHP003.Mimic,3) ,XIC(ControlLoop_FeedPumpAlarm.HIAlarm) XIO(ControlLoop_FeedPumpAlarm.HIHIAlarm) ] MOV(1,SIC001.DriveAlarmStatus) ,[LIM(4,SIC003DF.Mimic,5) ,LIM(4,DF3PHP003.Mimic,5) ,XIC(ControlLoop_FeedPumpAlarm.HIHIAlarm) ] MOV(2,SIC001.DriveAlarmStatus) ];
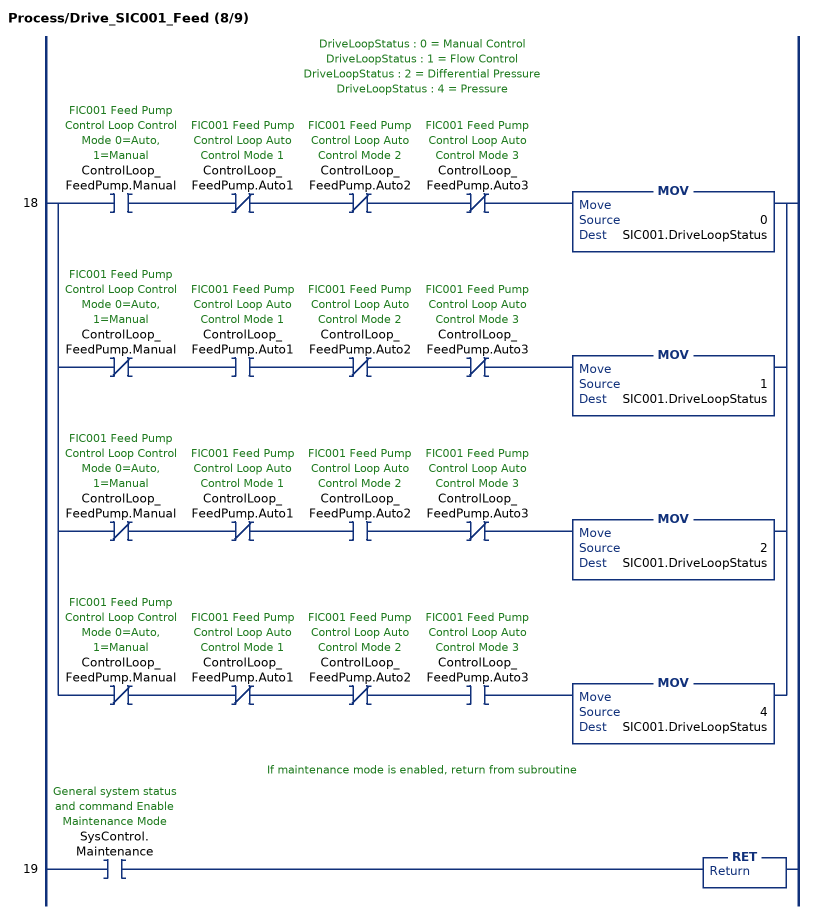
   // DriveLoopStatus : 0 = Manual Control
   //  DriveLoopStatus : 1 = Flow Control
   //  DriveLoopStatus : 2 = Differential Pressure
   //  DriveLoopStatus : 4 = Pressure
   18: [XIC(ControlLoop_FeedPump.Manual) XIO(ControlLoop_FeedPump.Auto1) XIO(ControlLoop_FeedPump.Auto2) XIO(ControlLoop_FeedPump.Auto3) MOV(0,SIC001.DriveLoopStatus) ,XIO(ControlLoop_FeedPump.Manual) XIC(ControlLoop_FeedPump.Auto1) XIO(ControlLoop_FeedPump.Auto2) XIO(ControlLoop_FeedPump.Auto3) MOV(1,SIC001.DriveLoopStatus) ,XIO(ControlLoop_FeedPump.Manual) XIO(ControlLoop_FeedPump.Auto1) XIC(ControlLoop_FeedPump.Auto2) XIO(ControlLoop_FeedPump.Auto3) MOV(2,SIC001.DriveLoopStatus) ,XIO(ControlLoop_FeedPump.Manual) XIO(ControlLoop_FeedPump.Auto1) XIO(ControlLoop_FeedPump.Auto2) XIC(ControlLoop_FeedPump.Auto3) MOV(4,SIC001.DriveLoopStatus) ];
   // If maintenance mode is enabled, return from subroutine
   19: XIC(SysControl.Maintenance)RET();
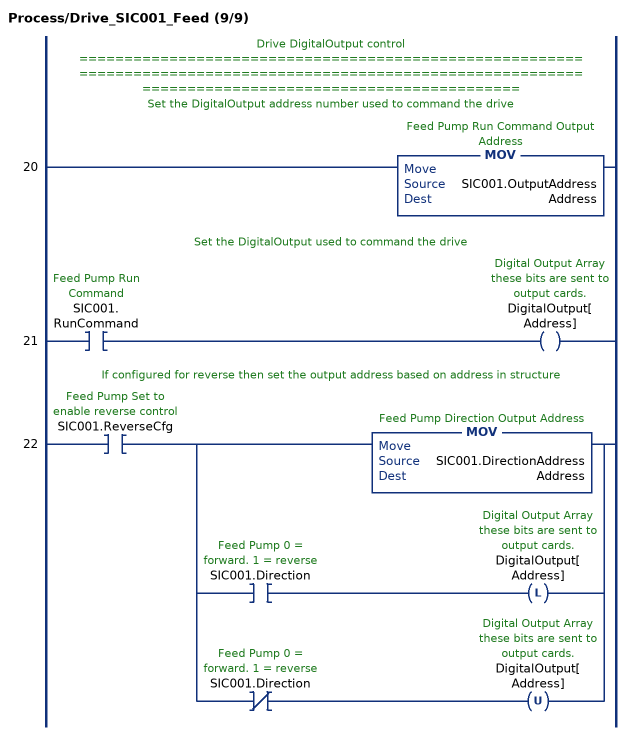
   // Drive DigitalOutput control
   // ==========================================================================================================================================================
   // Set the DigitalOutput address number used to command the drive
   20: MOV(SIC001.OutputAddress,Address);
   // Set the DigitalOutput used to command the drive
   21: XIC(SIC001.RunCommand)OTE(DigitalOutput[Address]);
   // If configured for reverse then set the output address based on address in structure
   22: XIC(SIC001.ReverseCfg)[MOV(SIC001.DirectionAddress,Address) ,XIC(SIC001.Direction) OTL(DigitalOutput[Address]) ,XIO(SIC001.Direction) OTU(DigitalOutput[Address]) ];
END_ROUTINE
